Fanuc KAREL source: kb00014.KL

-- PROVISIONAL review KL for V770-1; original PC SHA256 70427f56e2ad5cd1a681deb8bdb5189038b7071013c742739fd0b60e9270b5f9
-- Incomplete behavior may be omitted. Consult companion uncertainty JSON. Do not deploy.
PROGRAM KB00014
%NOLOCKGROUP
BEGIN
  -- UNRESOLVED_PC offsets 5-21; opcodes 27,22,31,23
  -- UNRESOLVED_PC offsets 26-30; opcodes 7F
END KB00014
